// TIA Portal V20 export
// export: Created 2026-10-20T18:55:52.7724836Z, ExportSetting None, DisplayName Totally Integrated Automation Portal, DisplayVersion V20 Update 6, DisplayName TIA Portal Openness, DisplayVersion V20 Update 6, DisplayName TIA Portal Version Control Interface, DisplayVersion V20 Update 6, DisplayName SINAMICS Startdrive Advanced, DisplayVersion V20 SP1, DisplayName SINAMICS Startdrive G130, G150, S120, S150, SINAMICS MV, G220, S200, S210, DisplayVersion V20 SP1, DisplayName SINAMICS Startdrive G110M, G120, G120C, G120D, G120P, G115D, DisplayVersion V20 SP1, DisplayName STEP 7 Professional, DisplayVersion V20 Update 6, DisplayName STEP 7 Safety, DisplayVersion V20 Update 2, DisplayName WinCC Basic/Comfort/Advanced, DisplayVersion V20 Update 6, DisplayName WinCC Unified, DisplayVersion V20 Update 6
VAR_GLOBAL   // PLC tag table "Lock_7"
   Lock_7_Estop_CH2 AT %I1806.3 : Bool;
   Lock_7_Estop_CH1 AT %I1806.2 : Bool;
   Lamps_7 AT %QB1491 : Byte;
   "Lock Reset_7" AT %Q1493.0 : Bool;
   "Solenoid Enable_7" AT %Q1492.0 : Bool;
   Lock_7_Closed_CH2 AT %I1806.1 : Bool;
   Switches_7 AT %IB1343 : Byte;
   Lock_7_Closed_CH1 AT %I1806.0 : Bool;
   Lock_7_Reset_Input2 AT %Q1807.1 : Bool;
   Lock_7_Reset_Input4 AT %Q1807.3 : Bool;
   Lock_7_Reset_Input3 AT %Q1807.2 : Bool;
   Lock_7_Reset_Input1 AT %Q1807.0 : Bool;
   "Lock Position_7" AT %I1345.0 : Bool;
   "Guard Position_7" AT %I1344.0 : Bool;
END_VAR
